FUNCTION_BLOCK FB_AliasLevel1
VAR
    {attribute 'pytmc' := '
        pv:LEVEL1
    '}
    stAlias : ST_Alias;

    {attribute 'pytmc' := '
        pv: LEVEL2
    '}
    fbAliasLevel2 : FB_AliasLevel2;
END_VAR

END_FUNCTION_BLOCK

(* stored: Version 1.1.0.1
   POU FB_AliasLevel1: Id {6270e95f-877e-47b3-8959-6bba924daa23}, SpecialFunc None *)
